// TIA Portal V17 export
// export: Created 2026-11-10T15:00:48.6641979Z, ExportSetting WithDefaults, DisplayName Totally Integrated Automation Portal, DisplayVersion V17, DisplayName TIA Portal Openness, DisplayVersion V17, DisplayName TIA Portal Version Control Interface, DisplayVersion V17, DisplayName STEP 7 Professional, DisplayVersion V17, DisplayName STEP 7 Safety, DisplayVersion V17, DisplayName WinCC Advanced, DisplayVersion V17
GraphicList "TruckFrames"  ListRange=Decimal, Mode=Simple
  GraphicListEntry   EntryType=Range, Picture=Truck_0
  GraphicListEntry   EntryType=Range, From=1, To=1, Picture=Truck_1
  GraphicListEntry   EntryType=Range, From=2, To=2, Picture=Truck_2
  GraphicListEntry   EntryType=Range, From=3, To=3, Picture=Truck_3
  GraphicListEntry   EntryType=Range, From=4, To=4, Picture=Truck_4
  GraphicListEntry   EntryType=Range, From=5, To=5, Picture=Truck_5
  GraphicListEntry   EntryType=Range, From=6, To=6, Picture=Truck_6
  GraphicListEntry   EntryType=Range, From=7, To=7, Picture=Truck_7
  GraphicListEntry   EntryType=Range, From=8, To=8, Picture=Truck_8
  GraphicListEntry   EntryType=Range, From=9, To=9, Picture=Truck_9
  GraphicListEntry   EntryType=Range, From=10, To=10, Picture=Truck_10
